INTERFACE ITcoComponent EXTENDS ITcoObject,ITcoRestorable, ITcoServiceable

END_INTERFACE

(* stored: Version 1.1.0.1
   Itf ITcoComponent: Id {ad6fdf47-e58a-0ffd-120f-617d765bd842} *)
